(* IEC 61131-3 sources: voltrus-explorers/crates/mt-plc-cli/tests/fixtures/fbd, 4 files *)

(* ---- counter.golden.st ---- *)
PROGRAM Counter
VAR_INPUT
    X0 : BOOL;
    X1 : BOOL;
END_VAR
VAR_OUTPUT
    Y0 : BOOL;
END_VAR
VAR
    part_counter : CTU;
END_VAR

    part_counter(CU := X0, R := X1, PV := 10);
    Y0 := part_counter.Q;
END_PROGRAM

(* ---- motor-start-stop.golden.st ---- *)
PROGRAM MotorStartStop
VAR_INPUT
    M0 : BOOL;
    X0 : BOOL;
    X1 : BOOL;
END_VAR
VAR_OUTPUT
    Y0 : BOOL;
END_VAR
VAR
    __t1 : BOOL;
END_VAR

    __t1 := X0 OR M0;
    Y0 := __t1 AND X1;
END_PROGRAM

(* ---- threshold-alarm.golden.st ---- *)
PROGRAM ThresholdAlarm
VAR_INPUT
    D0 : INT;
    D1 : INT;
END_VAR
VAR_OUTPUT
    Y0 : BOOL;
END_VAR
VAR
    __t1 : INT;
END_VAR

    __t1 := D0 + D1;
    Y0 := __t1 > 100;
END_PROGRAM

(* ---- timer-delay.golden.st ---- *)
PROGRAM TimerDelay
VAR_INPUT
    X0 : BOOL;
END_VAR
VAR_OUTPUT
    Y0 : BOOL;
END_VAR
VAR
    delay_timer : TON;
END_VAR

    delay_timer(IN := X0, PT := T#500MS);
    Y0 := delay_timer.Q;
END_PROGRAM
